INTERFACE I_Motor

METHOD M_Start : BOOL
VAR_INPUT
fSpeed:LREAL;
END_VAR
END_METHOD

PROPERTY P_State : E_MotorState
GET // PUBLIC
END_GET
END_PROPERTY

END_INTERFACE

(* stored: Version 1.1.0.1
   Itf I_Motor: Id {46ff3029-b598-47d7-91a3-580cfc33a5b0}
   Method M_Start: Id {46ed1309-6ee5-4a37-9839-e7ceecc70927}
   Property P_State: Id {1b52d863-ac8a-4690-b53b-de27d0ef148b}
   Get Get: Id {eff680a6-b354-44ae-8072-e9d624e8289b} *)
